Fanuc KAREL source: kt00133.KL

-- PROVISIONAL review KL for V940-1; original PC SHA256 f11f7a056740b2663708a1758b23eb1285db4e3de4100219be759173b954dab9
-- Incomplete behavior may be omitted. Consult companion uncertainty JSON. Do not deploy.
PROGRAM KT00133
%NOLOCKGROUP
VAR
  I1 : INTEGER
  OUT : INTEGER
-- UNRESOLVED_DECL Y2 type=002018
BEGIN
  -- V9_ZERO_TABLE_METADATA_HINT layout=0001; no indexed target words; source/name/runtime held
  -- UNRESOLVED_PC offsets 5-16; opcodes 2E,23
  -- UNRESOLVED_PC offsets 21-35; opcodes 2E,22,9D,33,B2
  -- UNRESOLVED_PC offsets 40-62; opcodes 21,22,9D,33,B1,55,23
  -- UNRESOLVED_PC offsets 67-71; opcodes 7F
END KT00133
